(* IEC 61131-3 sources: SRCI_CLIENT_PLC/RobotLibrary/Library/POUs/Calculation/MC_CalculateCartesianPosition/Structures, 4 files *)

(* ---- CalculateCartesianPositionOutCmd.st ---- *)
{attribute 'pack_mode' := '1'}
// -------------------------------------------------------------------------
//  SRCI Robot Library
// -------------------------------------------------------------------------
//
//  Object:      CalculateCartesianPositionOutCmd
//  Author:      Thorsten Brach
//  Date:        2024-06-05
//
//  Description:
//
//
//  Copyright:
//    (C) 2024 Thorsten Brach. All rights reserved
//             Licensed under the MIT License.
//
//  Disclaimer:
//    This project is provided without any guarantee and can be used for
//    private and commercial purposes. Any use is at the user’s
//    own risk and responsibility.
//
// -------------------------------------------------------------------------
TYPE CalculateCartesianPositionOutCmd :
STRUCT
  /// Index of target tool
  /// • 0: Flange (default)
  /// • 1..254: Tool frames
  TargetToolNoReturn       : USINT;
  /// Index of target frame
  /// •      0: WCS
  /// • 1..254: User frames
  TargetFrameNoReturn      : USINT;
  /// Calculated cartesian position
  CartesianPositionReturn  : RobotCartesianPosition;
END_STRUCT
END_TYPE

(* ---- CalculateCartesianPositionParCmd.st ---- *)
{attribute 'pack_mode' := '1'}
// -------------------------------------------------------------------------
//  SRCI Robot Library
// -------------------------------------------------------------------------
//
//  Object:      CalculateCartesianPositionParCmd
//  Author:      Thorsten Brach
//  Date:        2024-06-05
//
//  Description:
//
//
//  Copyright:
//    (C) 2024 Thorsten Brach. All rights reserved
//             Licensed under the MIT License.
//
//  Disclaimer:
//    This project is provided without any guarantee and can be used for
//    private and commercial purposes. Any use is at the user’s
//    own risk and responsibility.
//
// -------------------------------------------------------------------------
TYPE CalculateCartesianPositionParCmd :
STRUCT
  /// Index of initial frame
  /// • 0: WCS (default)
  /// • 1..254: User frames
  FrameNo            : USINT;
  /// Index of target frame
  /// • 0: WCS (default)
  /// • 1..254: User frames
  TargetFrameNo      : USINT;
  /// Robot cartesian position.
  CartesianPosition  : RobotCartesianPosition;
END_STRUCT
END_TYPE

(* ---- CalculateCartesianPositionRecvData.st ---- *)
{attribute 'pack_mode' := '1'}
// -------------------------------------------------------------------------
//  SRCI Robot Library
// -------------------------------------------------------------------------
//
//  Object:      CalculateCartesianPositionRecvData
//  Author:      Thorsten Brach
//  Date:        2024-06-05
//
//  Description:
//
//
//  Copyright:
//    (C) 2024 Thorsten Brach. All rights reserved
//             Licensed under the MIT License.
//
//  Disclaimer:
//    This project is provided without any guarantee and can be used for
//    private and commercial purposes. Any use is at the user’s
//    own risk and responsibility.
//
// -------------------------------------------------------------------------
TYPE CalculateCartesianPositionRecvData EXTENDS RspHeader :
STRUCT
  /// Index of target tool
  /// • 0: Flange (default)
  /// • 1..254: Tool frames
  TargetToolNoReturn       : USINT;
  /// Index of target frame
  /// •      0: WCS
  /// • 1..254: User frames
  TargetFrameNoReturn      : USINT;
  /// Calculated cartesian position
  CartesianPositionReturn  : RobotCartesianPosition;
END_STRUCT
END_TYPE

(* ---- CalculateCartesianPositionSendData.st ---- *)
{attribute 'pack_mode' := '1'}
// -------------------------------------------------------------------------
//  SRCI Robot Library
// -------------------------------------------------------------------------
//
//  Object:      CalculateCartesianPositionSendData
//  Author:      Thorsten Brach
//  Date:        2024-06-05
//
//  Description:
//
//
//  Copyright:
//    (C) 2024 Thorsten Brach. All rights reserved
//             Licensed under the MIT License.
//
//  Disclaimer:
//    This project is provided without any guarantee and can be used for
//    private and commercial purposes. Any use is at the user’s
//    own risk and responsibility.
//
// -------------------------------------------------------------------------
TYPE CalculateCartesianPositionSendData EXTENDS CmdHeader:
STRUCT
  /// Index of source frame
  /// • 0: WCS (default)
  /// • 1..254: User frames
  FrameNo           : USINT;
  /// Index of target frame
  /// • 0: WCS (default)
  /// • 1..254: User frames
  TargetFrameNo     : USINT;
  /// Robot cartesian position.
  CartesianPosition : RobotCartesianPosition;
END_STRUCT
END_TYPE
